(* Schneider Machine Expert - Basic project Gas_controller, file version 3.0.0.0 *)
(* ProjectInformations: Name=t-New project *)

HARDWARE
  Cpu 0: TM221ME16R/G
  ModuleExtensionObject 0: TM3AQ2/G
  EthernetConfiguration: NetworkName=M221, IpAllocationMode=FixedAddress, IpAddress=192.168.1.22, SubnetMask=255.255.255.0
  SerialLineConfiguration: Baud=Baud19200, Parity=ParityEven, DataBits=DataBits8, StopBits=StopBits1, PhysicalMedium=PhysicalMediumRs485, TransmissionMode=TransmissionModeModbusRtu, SlaveId=1, Addressing=SlaveAddressing
  MastTask: UsePeriodScanMode=false, PeriodScan=100
  FastTask: Period=255
  CpuBehavior: StartingMode=StartAsPreviousState, AutoSaveRamOnEeprom=true, WatchdogPeriod=250

SYMBOLS  (address, symbol, comment, settings)
  %S13      SB_FIRSTRUN  "Indicates the first controller cycle in RUN mode"
  %TM0        [Preset=20, Base=OneHundredMilliSeconds]
  %TM1        [Preset=600, Base=OneHundredMilliSeconds]
  %TM2        [Preset=10, Base=OneHundredMilliSeconds]
  %IW0.0      [Type=Type_0_10V, Scope=Scope_Normal, Minimum=0, Maximum=1000]
  %QW1.0      [Type=Type_4_20mA, Scope=Scope_Customized, Minimum=0, Maximum=10000]

POU t-New POU
  (* SectionNumber=1 *)

// Rung 0
  LD %S13                 (* SB_FIRSTRUN *)
  [ %MW0 := 0 ]
  [ %MW2 := 0 ]
  // as ST:
  //   IF SB_FIRSTRUN THEN %MW0 := 0; END_IF;
  //   IF SB_FIRSTRUN THEN %MW2 := 0; END_IF;

// Rung 1
  LD [ %MW1 <> %MW3 ]
  ST %M0
  // as ST:
  //   %M0 := %MW1 <> %MW3;

// Rung 2
  LD %M0
  [ %MW3 := %MW1 ]
  // as ST:
  //   IF %M0 THEN %MW3 := %MW1; END_IF;

// Rung 3
  BLK %TM0
  LDN %M0
  IN
  OUT_BLK
  LD Q
  ST %M1
  END_BLK
  // as ST:
  //   %TM0(IN := NOT %M0);
  //   %M1 := %TM0.Q;

// Rung 4
  LD %M1
  OR [ %MW2 <> 1 ]
  ST %M2
  // as ST:
  //   %M2 := %M1 OR %MW2 <> 1;

// Rung 5
  LDN %M2
  [ %MW10 := %MW0 ]
  // as ST:
  //   IF NOT %M2 THEN %MW10 := %MW0; END_IF;

// Rung 6
  LD %M2
  [ %MW10 := 0 ]
  // as ST:
  //   IF %M2 THEN %MW10 := 0; END_IF;

// Rung 7
  LD [ %MW10 > 10000 ]
  [ %MW10 := 10000 ]
  // as ST:
  //   IF %MW10 > 10000 THEN %MW10 := 10000; END_IF;

// Rung 8
  LD [ %MW10 < 0 ]
  [ %MW10 := 0 ]
  // as ST:
  //   IF %MW10 < 0 THEN %MW10 := 0; END_IF;

// Rung 9
  LDN %M100
  [ %QW1.0 := %MW10 ]
  // as ST:
  //   IF NOT %M100 THEN %QW1.0 := %MW10; END_IF;

// Rung 10
  LDN %M100
  [ %MW11 := %IW0.0 ]
  // as ST:
  //   IF NOT %M100 THEN %MW11 := %IW0.0; END_IF;

// Rung 11
  LDN %M100
  [ %MW12 := %MW11 - 200 ]
  [ %MW12 := %MW12 * 25 ]
  [ %MW12 := %MW12 / 2 ]
  // as ST:
  //   IF NOT %M100 THEN %MW12 := %MW11 - 200; END_IF;
  //   IF NOT %M100 THEN %MW12 := %MW12 * 25; END_IF;
  //   IF NOT %M100 THEN %MW12 := %MW12 / 2; END_IF;

// Rung 12
  LD [ %MW12 < 0 ]
  [ %MW12 := 0 ]
  // as ST:
  //   IF %MW12 < 0 THEN %MW12 := 0; END_IF;

// Rung 13
  LD [ %MW12 > 10000 ]
  [ %MW12 := 10000 ]
  // as ST:
  //   IF %MW12 > 10000 THEN %MW12 := 10000; END_IF;

// Rung 14
  LDN %M100
  [ %MW14 := %MW10 - %MW12 ]
  // as ST:
  //   IF NOT %M100 THEN %MW14 := %MW10 - %MW12; END_IF;

// Rung 15
  LD [ %MW14 > 200 ]
  OR [ %MW14 < -200 ]
  ST %M3
  // as ST:
  //   %M3 := %MW14 > 200 OR %MW14 < -200;

// Rung 16
  BLK %TM1
  LD %M3
  ANDN %M6
  IN
  OUT_BLK
  LD Q
  ST %M4
  END_BLK
  // as ST:
  //   %TM1(IN := %M3 AND NOT %M6);
  //   %M4 := %TM1.Q;

// Rung 17
  LDN %M3
  ANDN %M6
  ST %M5
  // as ST:
  //   %M5 := NOT %M3 AND NOT %M6;

// Rung 18
  BLK %TM2
  LD [ %MW11 < 180 ]
  IN
  OUT_BLK
  LD Q
  ST %M6
  END_BLK
  // as ST:
  //   %TM2(IN := %MW11 < 180);
  //   %M6 := %TM2.Q;

// Rung 19
  LD %M1
  ST %MW13:X0
  // as ST:
  //   %MW13:X0 := %M1;

// Rung 20
  LD %M4
  ST %MW13:X1
  // as ST:
  //   %MW13:X1 := %M4;

// Rung 21
  LD %M6
  ST %MW13:X2
  // as ST:
  //   %MW13:X2 := %M6;

// Rung 22
  LD %M5
  ST %MW13:X3
  // as ST:
  //   %MW13:X3 := %M5;

// Rung 23
  LD %I0.0
  ST %MW13:X4
  // as ST:
  //   %MW13:X4 := %I0.0;

// Rung 24
  LD %I0.1
  ST %MW13:X5
  // as ST:
  //   %MW13:X5 := %I0.1;
